Fanuc KAREL source: kt00062.KL

-- PROVISIONAL review KL for V940-1; original PC SHA256 7c378d6a0e7ed85b26257218e8c80f90470632edb7feda1a984f72c58da6bca4
-- Incomplete behavior may be omitted. Consult companion uncertainty JSON. Do not deploy.
PROGRAM KT00062
%NOLOCKGROUP
VAR
  OUT : REAL
-- UNRESOLVED_DECL H1 type=002017
-- UNRESOLVED_DECL Y2 type=002018
BEGIN
  -- V9_ZERO_TABLE_METADATA_HINT layout=0001; no indexed target words; source/name/runtime held
  -- UNRESOLVED_PC offsets 5-19; opcodes 2E,22,9D,33,B4
  -- UNRESOLVED_PC offsets 24-38; opcodes 2E,22,9D,33,B2
  -- UNRESOLVED_PC offsets 43-69; opcodes 22,9D,33,B3,22,9D,33,B1,53,64,23
  -- UNRESOLVED_PC offsets 74-78; opcodes 7F
END KT00062
